(* IEC 61131-3 sources: kns-port-domestic/upstream/plc-process-lib/src/POUs/Util/F_RateLimitLr, 2 files *)

(* ---- F_RateLimitLr.decl.st ---- *)
// Назначение: шаг ограничителя скорости изменения с состоянием в LREAL — как F_RateLimit, но текущее
//             значение и результат LREAL: малое приращение (медленная рампа при коротком цикле, 0,003 %/с
//             при цикле 1 мс рядом с 70 %) не теряется округлением до REAL на каждом шаге. Цель и скорости —
//             REAL (входы и Cfg устройств). Скорость 0 (или меньше) — без ограничения. lrDt_s <= 0 или
//             rTarget не конечно — значение не меняется. Рампы FB_ControlValve и FB_MotorVfd (CV-14, VFD-13).
// Автор:      kr0nsch
// Версия:     0.1.0
// Документ:   docs/fb/Functions.md
FUNCTION F_RateLimitLr : LREAL
VAR_INPUT
    lrCurrent     : LREAL;   // текущее значение (результат прошлого шага)
    rTarget       : REAL;    // цель
    rRateUp_ups   : REAL;    // предел скорости роста, инж. ед./с; <= 0 — без ограничения
    rRateDown_ups : REAL;    // предел скорости спада, инж. ед./с; <= 0 — без ограничения
    lrDt_s        : LREAL;   // шаг времени, с
END_VAR
VAR
    lrTarget : LREAL;        // цель в LREAL
END_VAR

(* ---- F_RateLimitLr.impl.st ---- *)
lrTarget := REAL_TO_LREAL(rTarget);
IF lrDt_s <= 0.0 OR NOT F_IsFinite(rIn := rTarget) THEN
    // шага нет или цель — мусор: значение не меняется
    F_RateLimitLr := lrCurrent;
ELSIF lrTarget > lrCurrent AND rRateUp_ups > 0.0 THEN
    // рост, ограничен сверху
    F_RateLimitLr := MIN(lrTarget, lrCurrent + REAL_TO_LREAL(rRateUp_ups) * lrDt_s);
ELSIF lrTarget < lrCurrent AND rRateDown_ups > 0.0 THEN
    // спад, ограничен снизу
    F_RateLimitLr := MAX(lrTarget, lrCurrent - REAL_TO_LREAL(rRateDown_ups) * lrDt_s);
ELSE
    // цель достигнута, скорость не ограничена или текущее значение не число: сразу к цели
    F_RateLimitLr := lrTarget;
END_IF
